Fanuc KAREL source: KT00545.KL

PROGRAM KT00545
%NOLOCKGROUP
VAR
  P1: JOINTPOS
  P2: XYZWPREXT
  OUT: XYZWPR
BEGIN
    P2.Y = 2.0
  OUT = P1 : P2
END KT00545
